RESOURCE RES0 : EMB_RES_ECO
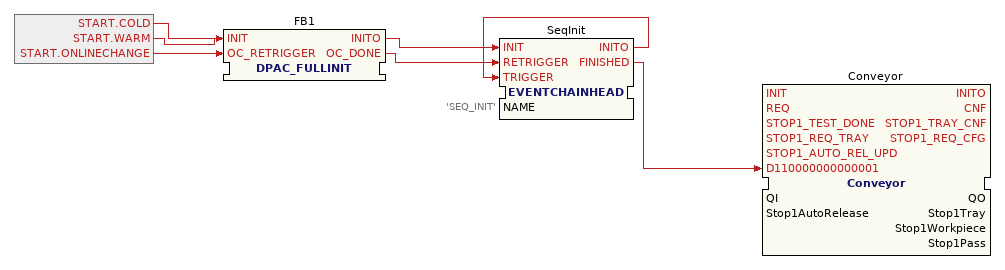
  FBS
    Conveyor : Conveyor;
    FB1 : DPAC_FULLINIT;
    SeqInit : EVENTCHAINHEAD(NAME := 'SEQ_INIT');
  END_FBS
  EVENT_CONNECTIONS
    START.COLD TO FB1.INIT;
    START.WARM TO FB1.INIT;
    START.ONLINECHANGE TO FB1.OC_RETRIGGER;
    FB1.INITO TO SeqInit.INIT;
    FB1.OC_DONE TO SeqInit.RETRIGGER;
    SeqInit.INITO TO SeqInit.TRIGGER;
    SeqInit.FINISHED TO Conveyor.D110000000000001;
  END_CONNECTIONS
END_RESOURCE
